DATA_BLOCK "TankA"
{ S7_Optimized_Access := 'TRUE' }
VERSION : 0.1
NON_RETAIN
"Tank"

BEGIN

END_DATA_BLOCK
